{attribute 'no_assign'}
FUNCTION_BLOCK FB_DO_WTURBINE_LD0_LPHD1_PhyNam EXTENDS FB_AcsiCommonDataClass
VAR_INPUT
	vendor: FB_AcsiDATypeVisString255 := (Fc:=ACSI_FC_DC, bLinkResult:=THIS^.AddDataToContainer(ipData:=vendor));
END_VAR
VAR
END_VAR

END_FUNCTION_BLOCK

(* stored: Version 1.1.0.1
   POU FB_DO_WTURBINE_LD0_LPHD1_PhyNam: Id {e55a5fe3-d98d-488b-8701-306d56fb9b9c}, SpecialFunc None *)
